// TIA Portal V21 export
// export: Created 2026-11-21T10:55:36.0366743Z, ExportSetting WithDefaults, DisplayName Totally Integrated Automation Portal, DisplayVersion V21, DisplayName STEP 7 Professional, DisplayVersion V21, DisplayName STEP 7 Safety, DisplayVersion V21, DisplayName Tech WebApplication, DisplayVersion V21, DisplayName WinCC Basic/Comfort/Advanced, DisplayVersion V21, DisplayName WinCC Unified, DisplayVersion V21
VAR_GLOBAL   // PLC tag table "Operator"
   Recipe_Selected AT %MW10 : Int;   // Recipe chosen on the panel, 1 to 3
   Bottles_Filled AT %MD12 : DInt;   // Bottles filled since the last start
END_VAR
